(* PLC project Machine_Expert_ Template, Machine Expert Logic Builder V19.2.3.0, author HP *)
(* stored: creationDateTime 2025-12-30T20:01:45.2018299, version 0.0.0.0, modificationDateTime 2025-12-30T20:01:00.7712215 *)

PROGRAM POU_Ladder
  VAR
    emergency_pb AT %IX0.0 : BOOL;
    System_ready AT %M?0 : BOOL;
    Input_1 AT %IX0.1 : BOOL;
    Output_1 AT %QX0.0 : BOOL;
  END_VAR
  VAR
    TON_0 : TON;
  END_VAR

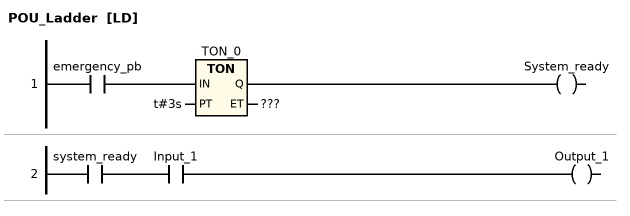
(* LD diagram, written out as Structured Text *)

TON_0(IN := emergency_pb, PT := t#3s, ET => ???);
System_ready := TON_0.Q;

Output_1 := system_ready AND Input_1;
END_PROGRAM
